// TIA Portal V20 export
TYPE "Kistler EO"
   STRUCT
      "X max" : Real;
      "X min" : Real;
      "Y max" : Real;
      "Y min" : Real;
      "EO Type" : USInt := 4;
      "EO Show Info" : Bool;
   END_STRUCT;
END_TYPE
